// TIA Portal V21 export
FUNCTION_BLOCK "LadBoxes"   // FB11, LAD
TITLE = Boxes
{ S7_Optimized_Access := 'TRUE' }
// Boxes in ladder: move, compare, add, timers, a counter and calls.
   VAR_INPUT
      level : Int;
      count : Bool;
      reset : Bool;
   END_VAR
   VAR_OUTPUT
      high : Bool;
      clamped : Int;
      done : Bool;
      pulse : Bool;
   END_VAR
   VAR
      delay : TON_TIME;
      "counter" : CTU_INT;
      pulser : "Pulse";
      copy : Int;
      sum : Int;
   END_VAR
BEGIN

REGION Network 1: Move
   // Copies the level.
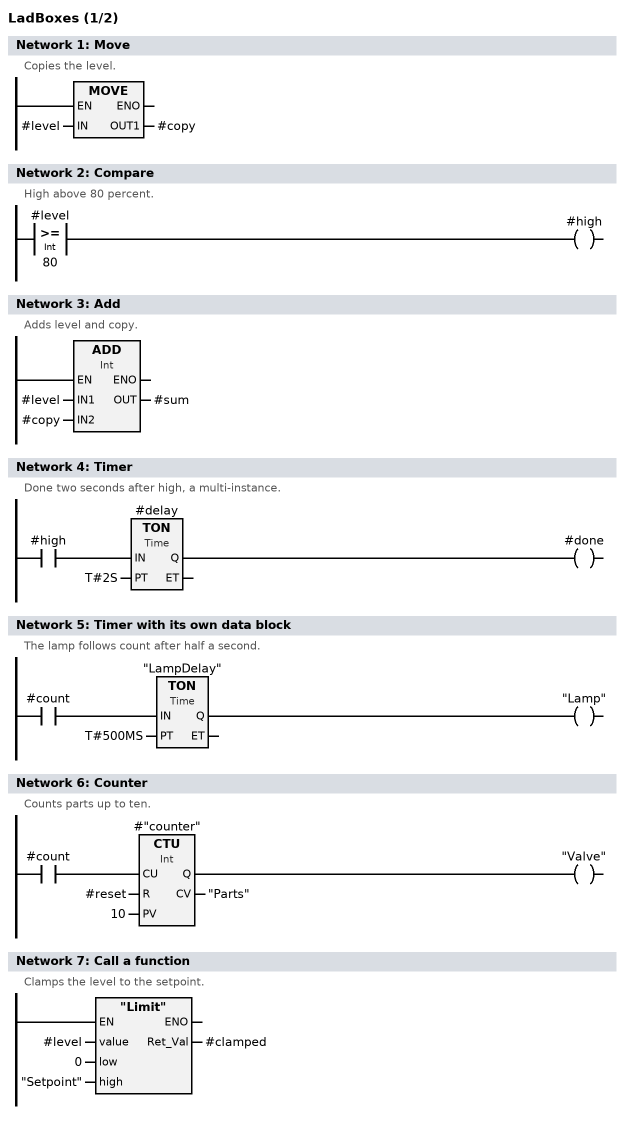
   RUNG wire#powerrail
      { S7_GenerateENO := "TRUE" } Move(in := #level, out1 => #copy)
   END_RUNG
   // the same network as SCL:
   #copy := #level;
END_REGION

REGION Network 2: Compare
   // High above 80 percent.
   RUNG wire#powerrail
      { S7_Templates := "SrcType := Int" } GE_Contact(in1 := #level, in2 := 80)
      Coil( #high )
   END_RUNG
   // the same network as SCL:
   #high := #level >= 80;
END_REGION

REGION Network 3: Add
   // Adds level and copy.
   RUNG wire#powerrail
      { S7_Templates := "SrcType := Int"; S7_GenerateENO := "TRUE" } Add(in1 := #level, in2 := #copy, out => #sum)
   END_RUNG
   // the same network as SCL:
   #sum := #level + #copy;
END_REGION

REGION Network 4: Timer
   // Done two seconds after high, a multi-instance.
   #delay(IN := #high, PT := T#2S);   // TON
   #done := #delay.Q;
END_REGION

REGION Network 5: Timer with its own data block
   // The lamp follows count after half a second.
   "LampDelay".TON(IN := #count, PT := T#500MS);
   "Lamp" := "LampDelay".Q;
END_REGION

REGION Network 6: Counter
   // Counts parts up to ten.
   #"counter"(CU := #count, R := #reset, PV := 10, CV => "Parts");   // CTU
   "Valve" := #"counter".Q;
END_REGION

REGION Network 7: Call a function
   // Clamps the level to the setpoint.
   RUNG wire#powerrail
      "Limit"(value := #level, low := 0, high := "Setpoint", Ret_Val => #clamped)
   END_RUNG
   // the same network as SCL:
   #clamped := "Limit"(value := #level, low := 0, high := "Setpoint");
END_REGION

REGION Network 8: Call a function block
   // A pulse on each count, a multi-instance.
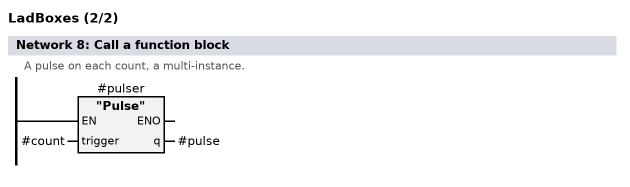
   RUNG wire#powerrail
      #pulser(trigger := #count, q => #pulse)
   END_RUNG
   // the same network as SCL:
   #pulser(trigger := #count, q => #pulse);   // "Pulse"
END_REGION
END_FUNCTION_BLOCK
